{attribute 'qualified_only'}
{attribute 'strict'}
{attribute 'to_string'}
TYPE E_UInt :
(
	eOptionA := 0,
	eOptionB,
	eOptionC
) UINT;
END_TYPE

(* stored: Version 1.1.0.1, ProductVersion 3.1.4026.19
   DUT E_UInt: Id {572f10bb-cda8-469d-a88f-30d25c2c08c7} *)
